// SIMATIC S7-200 project (STEP 7-Micro/WIN), CPU 226 CN REL 02.01

SYMBOL_TABLE USUARIO1
SI1              I0.0     // Sensor de riel
FCI              I0.1     // Final de carrera derecha
FCF              I0.2     // Final de carrera izquierda
QS               I2.6     // Zeta de emergencia
SB_1             I2.5     // Pulsador de marcha
SB_2             I2.4     // Pulsador de parada
SA               I2.7     // Selector de modo
PULSO            Q0.0     // Pulso
DIR              Q0.1     // Direccion
                 Q0.3     // Cilndro neumatico vertical
                 Q0.4     // Cilindro rotarorio anti horario
                 Q0.5     // Cilindro rotatorio horario
                 Q0.6     // Cilindro horizontal
                 Q0.7     // Garra cerrada
                 Q1.0     // Garra abierta
HL1              Q1.5     // Piloto Amarillo
HL2              Q1.6     // Piloto Verde
HL3              Q1.7     // Piloto Rojo
Mov1             V140.0   // primer movimiento
Mov2             V140.1   // segundo movimiento
END_SYMBOL_TABLE

ORGANIZATION_BLOCK PRINCIPAL:OB1
TITLE=COMENTARIOS DEL PROGRAMA
BEGIN
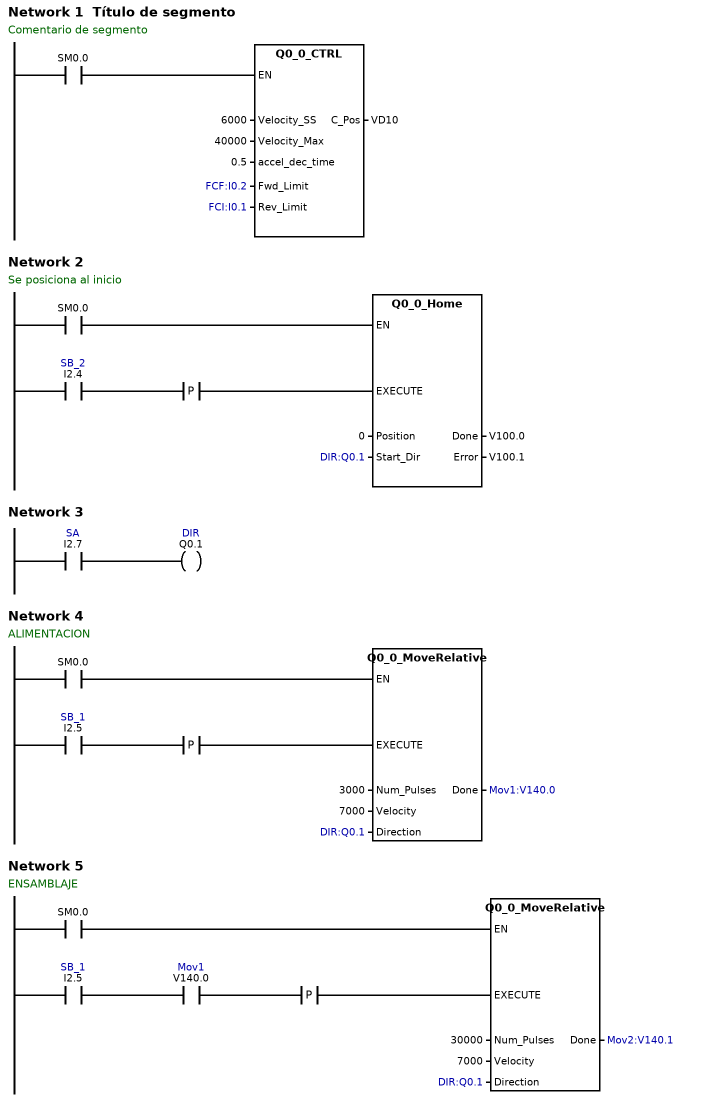
Network 1 // Título de segmento
// Comentario de segmento
LD     SM0.0
CALL   Q0_0_CTRL:SBR1, 6000, 40000, 0.5, FCF:I0.2, FCI:I0.1, VD10
Network 2
// Se posiciona al inicio 
LD     SM0.0
=      L60.0
LD     SB_2:I2.4
EU
=      L63.7
LD     L60.0
CALL   Q0_0_Home:SBR3, L63.7, 0, DIR:Q0.1, V100.0, V100.1
Network 3
LD     SA:I2.7
=      DIR:Q0.1
Network 4
// ALIMENTACION
LD     SM0.0
=      L60.0
LD     SB_1:I2.5
EU
=      L63.7
LD     L60.0
CALL   Q0_0_MoveRelative:SBR4, L63.7, 3000, 7000, DIR:Q0.1, Mov1:V140.0
Network 5
// ENSAMBLAJE
LD     SM0.0
=      L60.0
LD     SB_1:I2.5
A      Mov1:V140.0
EU
=      L63.7
LD     L60.0
CALL   Q0_0_MoveRelative:SBR4, L63.7, 30000, 7000, DIR:Q0.1, Mov2:V140.1
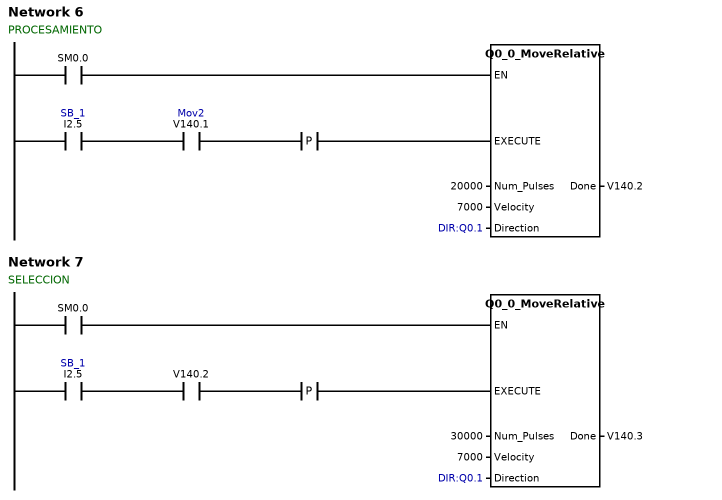
Network 6
// PROCESAMIENTO
LD     SM0.0
=      L60.0
LD     SB_1:I2.5
A      Mov2:V140.1
EU
=      L63.7
LD     L60.0
CALL   Q0_0_MoveRelative:SBR4, L63.7, 20000, 7000, DIR:Q0.1, V140.2
Network 7
// SELECCION
LD     SM0.0
=      L60.0
LD     SB_1:I2.5
A      V140.2
EU
=      L63.7
LD     L60.0
CALL   Q0_0_MoveRelative:SBR4, L63.7, 30000, 7000, DIR:Q0.1, V140.3
END_ORGANIZATION_BLOCK

// SBR1: protected block, not included

// SBR2: protected block, not included

// SBR3: protected block, not included

// SBR4: protected block, not included

// SBR5: protected block, not included
